TYPE ST_HeatUp :
STRUCT
	lrHeatUpForce						:LREAL;											(* HeatUp force [N] *)
	unHeatUpRamp						:UINT;											(* HeatUp ramp [s] *)
	unHeatUpTime						:UINT;											(* HeatUp time [s] *)
	lrVeloForceCtrlKp						:LREAL;											(* Velocity - force controller proportional band Kp *)
	lrVeloForceCtrlTi						:LREAL;											(* Velocity - force controller integral Ti *)
	lrVeloForceCtrlLimit					:LREAL;											(* Velocity - force controller limit  *)
END_STRUCT
END_TYPE

(* stored: Version 1.1.0.1, ProductVersion 3.1.4024.15
   DUT ST_HeatUp: Id {a07d18d1-c3e4-4401-892c-900351f2cca6} *)
